(* IEC 61131-3 sources: rusty/tests/lit/single/control_statements/case_unsigned_selector, 13 files *)

(* ---- alias_selector.st ---- *)
// RUN: %COMPILE %s && %RUN | %CHECK %s
//
// A selector whose type is an alias of USINT compares like a USINT in a CASE range.

TYPE Count : USINT; END_TYPE

FUNCTION classify : DINT
    VAR_INPUT
        x : Count;
    END_VAR
    CASE x OF
        11..254: classify := 1;
    ELSE
        classify := 0;
    END_CASE
END_FUNCTION

FUNCTION show
    VAR_INPUT
        x : Count;
    END_VAR
    printf('%u: %d$N', x, classify(x));
END_FUNCTION

FUNCTION main
    show(10);
    show(11);
    show(200);
    show(254);
    show(255);
    // CHECK:      10: 0
    // CHECK-NEXT: 11: 1
    // CHECK-NEXT: 200: 1
    // CHECK-NEXT: 254: 1
    // CHECK-NEXT: 255: 0
END_FUNCTION

(* ---- enum_selector_with_byte_base.st ---- *)
// RUN: %COMPILE %s && %RUN | %CHECK %s
//
// An enum with the unsigned base type BYTE compares as unsigned in a CASE range, so the range
// Low..Mid covers the variants 10 and 150 on both sides of the midpoint 128.

TYPE Level : (Low := 10, Mid := 150, High := 200) BYTE; END_TYPE

FUNCTION classify : DINT
    VAR_INPUT
        x : Level;
    END_VAR
    CASE x OF
        Low..Mid: classify := 1;
        High:     classify := 2;
    ELSE
        classify := 0;
    END_CASE
END_FUNCTION

FUNCTION main
    printf('Low: %d$N', classify(Low));
    printf('Mid: %d$N', classify(Mid));
    printf('High: %d$N', classify(High));
    // CHECK:      Low: 1
    // CHECK-NEXT: Mid: 1
    // CHECK-NEXT: High: 2
END_FUNCTION

(* ---- constant_range_bounds.st ---- *)
// RUN: %COMPILE %s && %RUN | %CHECK %s
//
// A range whose bounds are USINT constants compares like a range with literal bounds.

VAR_GLOBAL CONSTANT
    LOWER : USINT := 11;
    UPPER : USINT := 254;
END_VAR

FUNCTION classify : DINT
    VAR_INPUT
        x : USINT;
    END_VAR
    CASE x OF
        LOWER..UPPER: classify := 1;
    ELSE
        classify := 0;
    END_CASE
END_FUNCTION

FUNCTION show
    VAR_INPUT
        x : USINT;
    END_VAR
    printf('%u: %d$N', x, classify(x));
END_FUNCTION

FUNCTION main
    show(10);
    show(11);
    show(128);
    show(254);
    show(255);
    // CHECK:      10: 0
    // CHECK-NEXT: 11: 1
    // CHECK-NEXT: 128: 1
    // CHECK-NEXT: 254: 1
    // CHECK-NEXT: 255: 0
END_FUNCTION

(* ---- byte_range_around_midpoint.st ---- *)
// RUN: %COMPILE %s && %RUN | %CHECK %s
//
// A narrow range around the midpoint of a BYTE selector, 127..129, matches its three values and
// none of the neighbors.

FUNCTION classify : DINT
    VAR_INPUT
        x : BYTE;
    END_VAR
    CASE x OF
        127..129: classify := 1;
    ELSE
        classify := 0;
    END_CASE
END_FUNCTION

FUNCTION show
    VAR_INPUT
        x : BYTE;
    END_VAR
    printf('%u: %d$N', x, classify(x));
END_FUNCTION

FUNCTION main
    show(126);
    show(127);
    show(128);
    show(129);
    show(130);
    // CHECK:      126: 0
    // CHECK-NEXT: 127: 1
    // CHECK-NEXT: 128: 1
    // CHECK-NEXT: 129: 1
    // CHECK-NEXT: 130: 0
END_FUNCTION

(* ---- full_type_range.st ---- *)
// RUN: %COMPILE %s && %RUN | %CHECK %s
//
// A range over all values of a USINT selector, 0..255, matches every value, so ELSE never runs.

FUNCTION classify : DINT
    VAR_INPUT
        x : USINT;
    END_VAR
    CASE x OF
        0..255: classify := 1;
    ELSE
        classify := 0;
    END_CASE
END_FUNCTION

FUNCTION show
    VAR_INPUT
        x : USINT;
    END_VAR
    printf('%u: %d$N', x, classify(x));
END_FUNCTION

FUNCTION main
    show(0);
    show(127);
    show(128);
    show(255);
    // CHECK:      0: 1
    // CHECK-NEXT: 127: 1
    // CHECK-NEXT: 128: 1
    // CHECK-NEXT: 255: 1
END_FUNCTION

(* ---- range_in_label_list.st ---- *)
// RUN: %COMPILE %s && %RUN | %CHECK %s
//
// A label list that mixes single values and a range across the midpoint of a USINT selector
// matches all of them; the values that the list leaves out go to ELSE.

FUNCTION classify : DINT
    VAR_INPUT
        x : USINT;
    END_VAR
    CASE x OF
        0, 11..254, 255: classify := 1;
    ELSE
        classify := 0;
    END_CASE
END_FUNCTION

FUNCTION show
    VAR_INPUT
        x : USINT;
    END_VAR
    printf('%u: %d$N', x, classify(x));
END_FUNCTION

FUNCTION main
    show(0);
    show(10);
    show(11);
    show(200);
    show(255);
    // CHECK:      0: 1
    // CHECK-NEXT: 10: 0
    // CHECK-NEXT: 11: 1
    // CHECK-NEXT: 200: 1
    // CHECK-NEXT: 255: 1
END_FUNCTION

(* ---- ranges_in_lower_and_upper_half.st ---- *)
// RUN: %COMPILE %s && %RUN | %CHECK %s
//
// Ranges that stay in one half of a USINT selector split the values at the midpoint 128.

FUNCTION classify : DINT
    VAR_INPUT
        x : USINT;
    END_VAR
    CASE x OF
        0..127:   classify := 1;
        128..255: classify := 2;
    ELSE
        classify := 0;
    END_CASE
END_FUNCTION

FUNCTION show
    VAR_INPUT
        x : USINT;
    END_VAR
    printf('%u: %d$N', x, classify(x));
END_FUNCTION

FUNCTION main
    show(0);
    show(127);
    show(128);
    show(255);
    // CHECK:      0: 1
    // CHECK-NEXT: 127: 1
    // CHECK-NEXT: 128: 2
    // CHECK-NEXT: 255: 2
END_FUNCTION

(* ---- signed_range_across_zero.st ---- *)
// RUN: %COMPILE %s && %RUN | %CHECK %s
//
// A range on a signed SINT selector compares the selector as a signed value, so ranges with
// negative bounds and ranges across zero match as written.

FUNCTION classify : DINT
    VAR_INPUT
        x : SINT;
    END_VAR
    CASE x OF
        -128..-101: classify := 1;
        -100..100:  classify := 2;
    ELSE
        classify := 0;
    END_CASE
END_FUNCTION

FUNCTION show
    VAR_INPUT
        x : SINT;
    END_VAR
    printf('%d: %d$N', x, classify(x));
END_FUNCTION

FUNCTION main
    show(-128);
    show(-101);
    show(-100);
    show(0);
    show(100);
    show(101);
    show(127);
    // CHECK:      -128: 1
    // CHECK-NEXT: -101: 1
    // CHECK-NEXT: -100: 2
    // CHECK-NEXT: 0: 2
    // CHECK-NEXT: 100: 2
    // CHECK-NEXT: 101: 0
    // CHECK-NEXT: 127: 0
END_FUNCTION

(* ---- subrange_selector.st ---- *)
// RUN: %COMPILE %s && %RUN | %CHECK %s
//
// A selector whose type is a subrange of USINT compares like a USINT in a CASE range.

FUNCTION classify : DINT
    VAR_INPUT
        x : USINT(10..250);
    END_VAR
    CASE x OF
        100..200: classify := 1;
    ELSE
        classify := 0;
    END_CASE
END_FUNCTION

FUNCTION show
    VAR_INPUT
        x : USINT(10..250);
    END_VAR
    printf('%u: %d$N', x, classify(x));
END_FUNCTION

FUNCTION main
    show(99);
    show(100);
    show(150);
    show(200);
    show(201);
    // CHECK:      99: 0
    // CHECK-NEXT: 100: 1
    // CHECK-NEXT: 150: 1
    // CHECK-NEXT: 200: 1
    // CHECK-NEXT: 201: 0
END_FUNCTION

(* ---- udint_range_across_midpoint.st ---- *)
// RUN: %COMPILE %s && %RUN | %CHECK %s
//
// A range on a UDINT selector across the midpoint 2^31 matches every value between its bounds.

FUNCTION classify : DINT
    VAR_INPUT
        x : UDINT;
    END_VAR
    CASE x OF
        16#7FFF_FFFF..16#8000_0001: classify := 1;
    ELSE
        classify := 0;
    END_CASE
END_FUNCTION

FUNCTION show
    VAR_INPUT
        x : UDINT;
    END_VAR
    printf('%u: %d$N', x, classify(x));
END_FUNCTION

FUNCTION main
    show(16#7FFF_FFFE);
    show(16#7FFF_FFFF);
    show(16#8000_0000);
    show(16#8000_0001);
    show(16#8000_0002);
    // CHECK:      2147483646: 0
    // CHECK-NEXT: 2147483647: 1
    // CHECK-NEXT: 2147483648: 1
    // CHECK-NEXT: 2147483649: 1
    // CHECK-NEXT: 2147483650: 0
END_FUNCTION

(* ---- uint_range_across_midpoint.st ---- *)
// RUN: %COMPILE %s && %RUN | %CHECK %s
//
// A range on a UINT selector across the midpoint 32768 matches every value between its bounds.

FUNCTION classify : DINT
    VAR_INPUT
        x : UINT;
    END_VAR
    CASE x OF
        1..65534: classify := 1;
    ELSE
        classify := 0;
    END_CASE
END_FUNCTION

FUNCTION show
    VAR_INPUT
        x : UINT;
    END_VAR
    printf('%u: %d$N', x, classify(x));
END_FUNCTION

FUNCTION main
    show(0);
    show(1);
    show(32767);
    show(32768);
    show(65534);
    show(65535);
    // CHECK:      0: 0
    // CHECK-NEXT: 1: 1
    // CHECK-NEXT: 32767: 1
    // CHECK-NEXT: 32768: 1
    // CHECK-NEXT: 65534: 1
    // CHECK-NEXT: 65535: 0
END_FUNCTION

(* ---- ulint_range_across_midpoint.st ---- *)
// RUN: %COMPILE %s && %RUN | %CHECK %s
//
// A range on a ULINT selector across the midpoint 2^63 matches every value between its bounds.

FUNCTION classify : DINT
    VAR_INPUT
        x : ULINT;
    END_VAR
    CASE x OF
        16#7FFF_FFFF_FFFF_FFFF..16#8000_0000_0000_0001: classify := 1;
    ELSE
        classify := 0;
    END_CASE
END_FUNCTION

FUNCTION show
    VAR_INPUT
        x : ULINT;
    END_VAR
    printf('%llu: %d$N', x, classify(x));
END_FUNCTION

FUNCTION main
    show(16#7FFF_FFFF_FFFF_FFFE);
    show(16#7FFF_FFFF_FFFF_FFFF);
    show(16#8000_0000_0000_0000);
    show(16#8000_0000_0000_0001);
    show(16#8000_0000_0000_0002);
    // CHECK:      9223372036854775806: 0
    // CHECK-NEXT: 9223372036854775807: 1
    // CHECK-NEXT: 9223372036854775808: 1
    // CHECK-NEXT: 9223372036854775809: 1
    // CHECK-NEXT: 9223372036854775810: 0
END_FUNCTION

(* ---- usint_range_across_midpoint.st ---- *)
// RUN: %COMPILE %s && %RUN | %CHECK %s
//
// A range on a USINT selector whose bounds lie on both sides of the midpoint 128 matches every
// value between them. Single labels and ranges in the lower half keep working next to it.

FUNCTION classify : DINT
    VAR_INPUT
        x : USINT;
    END_VAR
    CASE x OF
        0:       classify := 1;
        1..9:    classify := 2;
        11..254: classify := 3;
        255:     classify := 4;
    END_CASE
END_FUNCTION

FUNCTION show
    VAR_INPUT
        x : USINT;
    END_VAR
    printf('%u: %d$N', x, classify(x));
END_FUNCTION

FUNCTION main
    show(0);
    show(9);
    show(10);
    show(11);
    show(127);
    show(128);
    show(254);
    show(255);
    // CHECK:      0: 1
    // CHECK-NEXT: 9: 2
    // CHECK-NEXT: 10: 0
    // CHECK-NEXT: 11: 3
    // CHECK-NEXT: 127: 3
    // CHECK-NEXT: 128: 3
    // CHECK-NEXT: 254: 3
    // CHECK-NEXT: 255: 4
END_FUNCTION
